// TIA Portal V20 export
FUNCTION_BLOCK "PR_UnloadingSeq_Soft2.0_workflow_f29f28"   // FB54, LAD
{ S7_Optimized_Access := 'TRUE' }
// stored: MemoryReserve 100, SetENOAutomatically false
   VAR_INPUT
      iAbort : Bool;
      iAutoRunning : Bool;
      iFaultReset : Bool;
      iGantryAtPick : Bool;
      iManualEntryConfirm : Bool;
      iPartPickOver : Bool;
      iPartPresent : Bool;
      iPickConfirmed : Bool;
      iRFIDReadError : Bool;
      iRFIDReadOver : Bool;
      iRFWriteDone : Bool;
      iRFWriteError : Bool;
      iRTR_Frm_Gantry : Bool;
      iReject : Bool;
      iReset_fault : Bool;
      iRetry : Bool;
      iRetryCount : Int;
      iSstMode : Bool;
      iSstPB : Bool;
      iStartFrmFibroSeq : Bool;
      iSystemAtHome : Bool;
      iUnloadGantryAtSafe : Bool;
   END_VAR
   VAR_OUTPUT
      qError : Array[0..2] of Bool;
      qMessage : Array[0..0] of Bool;
      qUnloadOver : Bool;
   END_VAR
   VAR
      c120_ChkPartAbsent_T1 : Bool;
      c120_ChkPartAbsent_T2 : Bool;
      c130_WtOpDecisionPick_T1 : Bool;
      c130_WtOpDecisionPick_T2 : Bool;
      c140_WtRFIDWriteOver_T1 : Bool;
      c140_WtRFIDWriteOver_T2 : Bool;
      c150_ChkRFWriteRetryCount_T1 : Bool;
      c150_ChkRFWriteRetryCount_T2 : Bool;
      c160_WtOpDecisionWrite_T1 : Bool;
      c160_WtOpDecisionWrite_T2 : Bool;
      c20_ChkRecoveryStatus_T1 : Bool;
      c20_ChkRecoveryStatus_T2 : Bool;
      c20_ChkRecoveryStatus_T3 : Bool;
      c50_WtRFIDReadOver_T1 : Bool;
      c50_WtRFIDReadOver_T2 : Bool;
      c60_ChkRetryCountOver_T1 : Bool;
      c60_ChkRetryCountOver_T2 : Bool;
      c70_WtOpDecisionRead_T1 : Bool;
      c70_WtOpDecisionRead_T2 : Bool;
      c80_ChkPartWorkable_T1 : Bool;
      c80_ChkPartWorkable_T2 : Bool;
      StateNo : Int;
      s100_WtGantryAtPick : Bool;
      s100_WtGantryAtPick_T1 : Bool;
      s10_WtStartFrmMain : Bool;
      s10_WtStartFrmMain_T1 : Bool;
      s110_WtPartPick : Bool;
      s110_WtPartPick_T1 : Bool;
      s120_ChkPartAbsent : Bool;
      s120_ChkPartAbsent_T1 : Bool;
      s120_ChkPartAbsent_T2 : Bool;
      s130_WtOpDecisionPick : Bool;
      s130_WtOpDecisionPick_T1 : Bool;
      s130_WtOpDecisionPick_T2 : Bool;
      s140_WtRFIDWriteOver : Bool;
      s140_WtRFIDWriteOver_T1 : Bool;
      s140_WtRFIDWriteOver_T2 : Bool;
      s150_ChkRFWriteRetryCount : Bool;
      s150_ChkRFWriteRetryCount_T1 : Bool;
      s150_ChkRFWriteRetryCount_T2 : Bool;
      s160_WtOpDecisionWrite : Bool;
      s160_WtOpDecisionWrite_T1 : Bool;
      s160_WtOpDecisionWrite_T2 : Bool;
      s170_ChkSystemAtHome : Bool;
      s170_ChkSystemAtHome_T1 : Bool;
      s180_WtStartLow : Bool;
      s180_WtStartLow_T1 : Bool;
      s1_WtResetReleased : Bool;
      s1_WtResetReleased_T1 : Bool;
      s20_ChkRecoveryStatus : Bool;
      s20_ChkRecoveryStatus_T1 : Bool;
      s20_ChkRecoveryStatus_T2 : Bool;
      s20_ChkRecoveryStatus_T3 : Bool;
      s30_WtOperatorAck : Bool;
      s30_WtOperatorAck_T1 : Bool;
      s40_WtAllAxesSafe : Bool;
      s40_WtAllAxesSafe_T1 : Bool;
      s50_WtRFIDReadOver : Bool;
      s50_WtRFIDReadOver_T1 : Bool;
      s50_WtRFIDReadOver_T2 : Bool;
      s60_ChkRetryCountOver : Bool;
      s60_ChkRetryCountOver_T1 : Bool;
      s60_ChkRetryCountOver_T2 : Bool;
      s70_WtOpDecisionRead : Bool;
      s70_WtOpDecisionRead_T1 : Bool;
      s70_WtOpDecisionRead_T2 : Bool;
      s80_ChkPartWorkable : Bool;
      s80_ChkPartWorkable_T1 : Bool;
      s80_ChkPartWorkable_T2 : Bool;
      s90_WtRTRFrmGantry : Bool;
      s90_WtRTRFrmGantry_T1 : Bool;
      sAbnormalStatus : Bool;
      sPartWorkable : Bool;
      sRFReadRetryCount : Int;
      sRFWriteRetryCount : Int;
      sSst : Bool;
      sSstPulse : Bool;
      sSstRise : Bool;
      sStWtResetRel : Bool;
      sStWtResetRel_T1 : Bool;
      sUnloadingActive : Bool;
   END_VAR
   VAR_TEMP
      tOne : Bool;
   END_VAR
   VAR_TEMP   // added for the SCL form of the ladder/FBD networks
      _w1 : Bool;
      _w2 : Bool;
   END_VAR
BEGIN

REGION Network 1
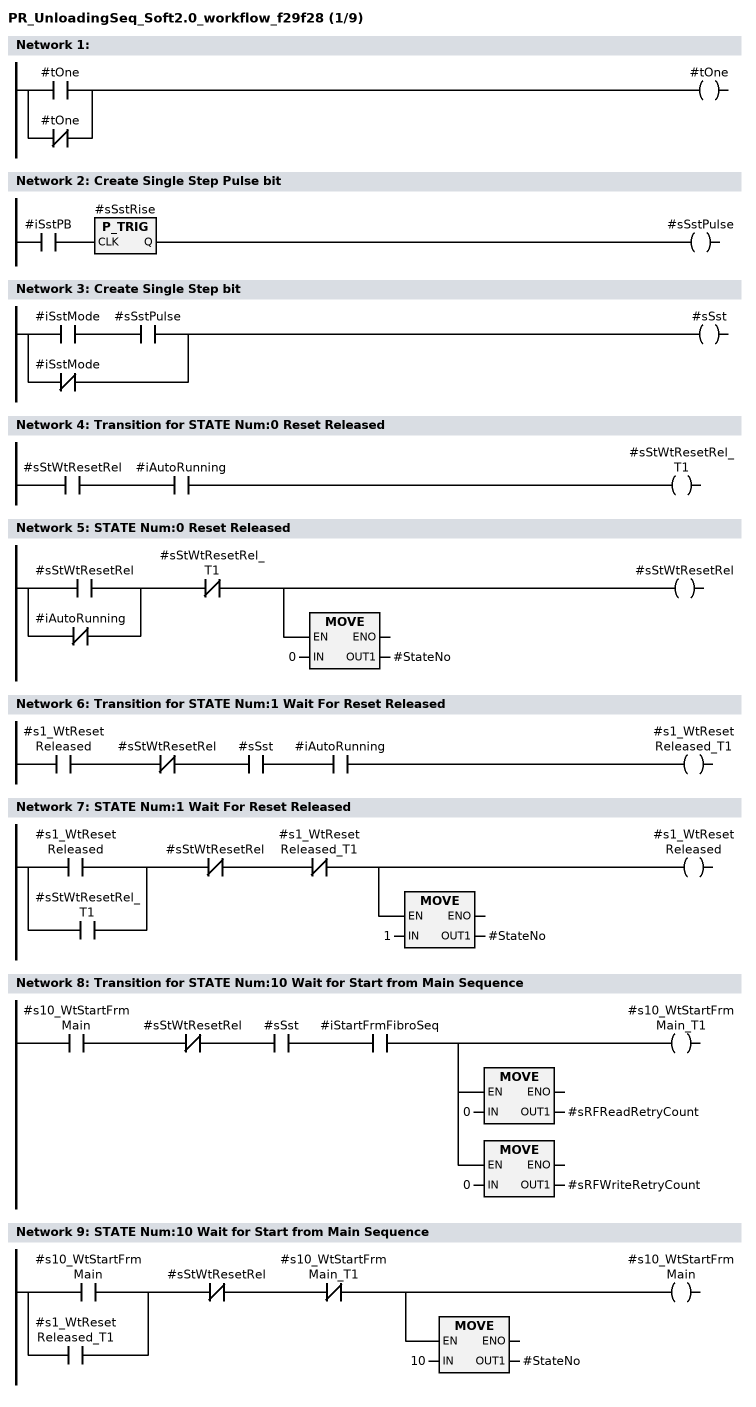
   RUNG wire#powerrail
      Contact( #tOne )
      wire#w1
      Coil( #tOne )
   END_RUNG
   RUNG wire#powerrail
      I_Contact( #tOne )
   END_RUNG wire#w1
   // the same network as SCL:
   #tOne := #tOne OR NOT #tOne;
END_REGION

REGION Network 2: Create Single Step Pulse bit
   RUNG wire#powerrail
      Contact( #iSstPB )
      P_Trig( #sSstRise )
      Coil( #sSstPulse )
   END_RUNG
   // the same network as SCL:
   #_w1 := #iSstPB AND NOT #sSstRise;   // rising edge
   #sSstRise := #iSstPB;
   #sSstPulse := #_w1;
END_REGION

REGION Network 3: Create Single Step bit
   RUNG wire#powerrail
      Contact( #iSstMode )
      Contact( #sSstPulse )
      wire#w1
      Coil( #sSst )
   END_RUNG
   RUNG wire#powerrail
      I_Contact( #iSstMode )
   END_RUNG wire#w1
   // the same network as SCL:
   #sSst := (#iSstMode AND #sSstPulse) OR NOT #iSstMode;
END_REGION

REGION Network 4: Transition for STATE Num:0 Reset Released
   RUNG wire#powerrail
      Contact( #sStWtResetRel )
      Contact( #iAutoRunning )
      Coil( #sStWtResetRel_T1 )
   END_RUNG
   // the same network as SCL:
   #sStWtResetRel_T1 := #sStWtResetRel AND #iAutoRunning;
END_REGION

REGION Network 5: STATE Num:0 Reset Released
   RUNG wire#powerrail
      Contact( #sStWtResetRel )
      wire#w1
      I_Contact( #sStWtResetRel_T1 )
      wire#w2
      Coil( #sStWtResetRel )
   END_RUNG
   RUNG wire#powerrail
      I_Contact( #iAutoRunning )
   END_RUNG wire#w1
   RUNG wire#w2
      { S7_GenerateENO := "TRUE" } Move(in := 0, out1 => #StateNo)
   END_RUNG
   // the same network as SCL:
   #sStWtResetRel := (#sStWtResetRel OR NOT #iAutoRunning) AND NOT #sStWtResetRel_T1;
   IF #sStWtResetRel THEN #StateNo := 0; END_IF;
END_REGION

REGION Network 6: Transition for STATE Num:1 Wait For Reset Released
   RUNG wire#powerrail
      Contact( #s1_WtResetReleased )
      I_Contact( #sStWtResetRel )
      Contact( #sSst )
      Contact( #iAutoRunning )
      Coil( #s1_WtResetReleased_T1 )
   END_RUNG
   // the same network as SCL:
   #s1_WtResetReleased_T1 := #s1_WtResetReleased AND NOT #sStWtResetRel AND #sSst AND #iAutoRunning;
END_REGION

REGION Network 7: STATE Num:1 Wait For Reset Released
   RUNG wire#powerrail
      Contact( #s1_WtResetReleased )
      wire#w1
      I_Contact( #sStWtResetRel )
      I_Contact( #s1_WtResetReleased_T1 )
      wire#w2
      Coil( #s1_WtResetReleased )
   END_RUNG
   RUNG wire#powerrail
      Contact( #sStWtResetRel_T1 )
   END_RUNG wire#w1
   RUNG wire#w2
      { S7_GenerateENO := "TRUE" } Move(in := 1, out1 => #StateNo)
   END_RUNG
   // the same network as SCL:
   #s1_WtResetReleased := (#s1_WtResetReleased OR #sStWtResetRel_T1) AND NOT #sStWtResetRel AND NOT #s1_WtResetReleased_T1;
   IF #s1_WtResetReleased THEN #StateNo := 1; END_IF;
END_REGION

REGION Network 8: Transition for STATE Num:10 Wait for Start from Main Sequence
   RUNG wire#powerrail
      Contact( #s10_WtStartFrmMain )
      I_Contact( #sStWtResetRel )
      Contact( #sSst )
      Contact( #iStartFrmFibroSeq )
      wire#w1
      Coil( #s10_WtStartFrmMain_T1 )
   END_RUNG
   RUNG wire#w1
      Move(in := 0, out1 => #sRFReadRetryCount)
   END_RUNG
   RUNG wire#w1
      Move(in := 0, out1 => #sRFWriteRetryCount)
   END_RUNG
   // the same network as SCL:
   #s10_WtStartFrmMain_T1 := #s10_WtStartFrmMain AND NOT #sStWtResetRel AND #sSst AND #iStartFrmFibroSeq;
   IF #s10_WtStartFrmMain_T1 THEN
       #sRFReadRetryCount := 0;
       #sRFWriteRetryCount := 0;
   END_IF;
END_REGION

REGION Network 9: STATE Num:10 Wait for Start from Main Sequence
   RUNG wire#powerrail
      Contact( #s10_WtStartFrmMain )
      wire#w1
      I_Contact( #sStWtResetRel )
      I_Contact( #s10_WtStartFrmMain_T1 )
      wire#w2
      Coil( #s10_WtStartFrmMain )
   END_RUNG
   RUNG wire#powerrail
      Contact( #s1_WtResetReleased_T1 )
   END_RUNG wire#w1
   RUNG wire#w2
      { S7_GenerateENO := "TRUE" } Move(in := 10, out1 => #StateNo)
   END_RUNG
   // the same network as SCL:
   #s10_WtStartFrmMain := (#s10_WtStartFrmMain OR #s1_WtResetReleased_T1) AND NOT #sStWtResetRel AND NOT #s10_WtStartFrmMain_T1;
   IF #s10_WtStartFrmMain THEN #StateNo := 10; END_IF;
END_REGION

REGION Network 10: Condition1 for STATE Num:20 Chek Recovery Status
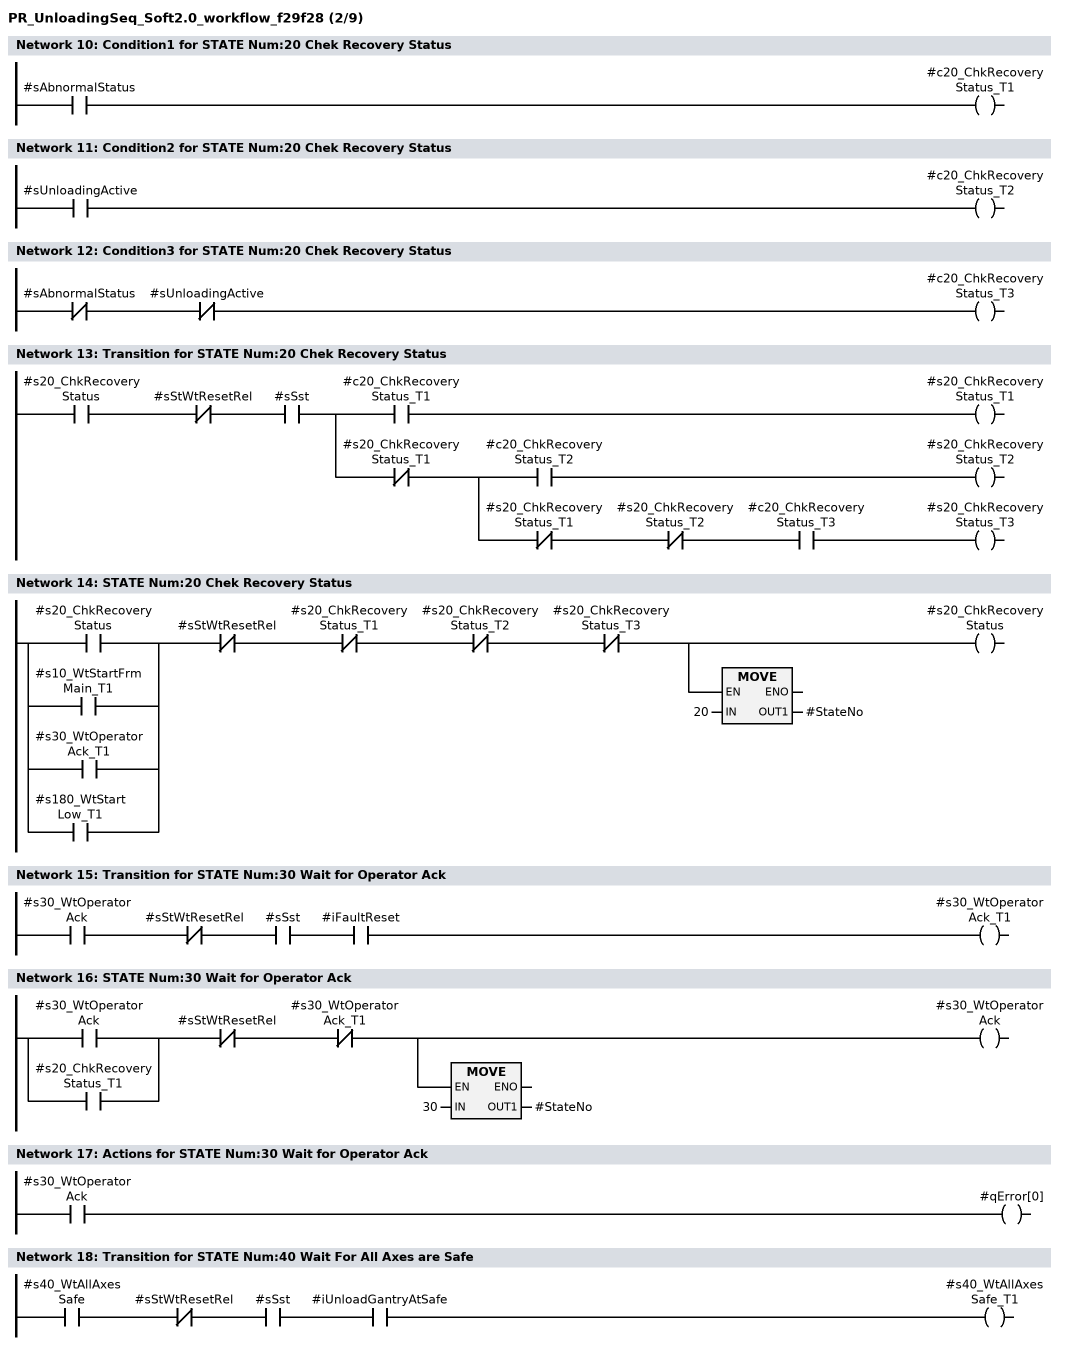
   RUNG wire#powerrail
      Contact( #sAbnormalStatus )
      Coil( #c20_ChkRecoveryStatus_T1 )
   END_RUNG
   // the same network as SCL:
   #c20_ChkRecoveryStatus_T1 := #sAbnormalStatus;
END_REGION

REGION Network 11: Condition2 for STATE Num:20 Chek Recovery Status
   RUNG wire#powerrail
      Contact( #sUnloadingActive )
      Coil( #c20_ChkRecoveryStatus_T2 )
   END_RUNG
   // the same network as SCL:
   #c20_ChkRecoveryStatus_T2 := #sUnloadingActive;
END_REGION

REGION Network 12: Condition3 for STATE Num:20 Chek Recovery Status
   RUNG wire#powerrail
      I_Contact( #sAbnormalStatus )
      I_Contact( #sUnloadingActive )
      Coil( #c20_ChkRecoveryStatus_T3 )
   END_RUNG
   // the same network as SCL:
   #c20_ChkRecoveryStatus_T3 := NOT #sAbnormalStatus AND NOT #sUnloadingActive;
END_REGION

REGION Network 13: Transition for STATE Num:20 Chek Recovery Status
   RUNG wire#powerrail
      Contact( #s20_ChkRecoveryStatus )
      I_Contact( #sStWtResetRel )
      Contact( #sSst )
      wire#w1
      Contact( #c20_ChkRecoveryStatus_T1 )
      Coil( #s20_ChkRecoveryStatus_T1 )
   END_RUNG
   RUNG wire#w1
      I_Contact( #s20_ChkRecoveryStatus_T1 )
      wire#w2
      Contact( #c20_ChkRecoveryStatus_T2 )
      Coil( #s20_ChkRecoveryStatus_T2 )
   END_RUNG
   RUNG wire#w2
      I_Contact( #s20_ChkRecoveryStatus_T1 )
      I_Contact( #s20_ChkRecoveryStatus_T2 )
      Contact( #c20_ChkRecoveryStatus_T3 )
      Coil( #s20_ChkRecoveryStatus_T3 )
   END_RUNG
   // the same network as SCL:
   #_w1 := #s20_ChkRecoveryStatus AND NOT #sStWtResetRel AND #sSst;
   #s20_ChkRecoveryStatus_T1 := #_w1 AND #c20_ChkRecoveryStatus_T1;
   #_w2 := #_w1 AND NOT #s20_ChkRecoveryStatus_T1;
   #s20_ChkRecoveryStatus_T2 := #_w2 AND #c20_ChkRecoveryStatus_T2;
   #s20_ChkRecoveryStatus_T3 := #_w2 AND NOT #s20_ChkRecoveryStatus_T1 AND NOT #s20_ChkRecoveryStatus_T2 AND #c20_ChkRecoveryStatus_T3;
END_REGION

REGION Network 14: STATE Num:20 Chek Recovery Status
   RUNG wire#powerrail
      Contact( #s20_ChkRecoveryStatus )
      wire#w1
      I_Contact( #sStWtResetRel )
      I_Contact( #s20_ChkRecoveryStatus_T1 )
      I_Contact( #s20_ChkRecoveryStatus_T2 )
      I_Contact( #s20_ChkRecoveryStatus_T3 )
      wire#w2
      Coil( #s20_ChkRecoveryStatus )
   END_RUNG
   RUNG wire#powerrail
      Contact( #s10_WtStartFrmMain_T1 )
   END_RUNG wire#w1
   RUNG wire#powerrail
      Contact( #s30_WtOperatorAck_T1 )
   END_RUNG wire#w1
   RUNG wire#powerrail
      Contact( #s180_WtStartLow_T1 )
   END_RUNG wire#w1
   RUNG wire#w2
      { S7_GenerateENO := "TRUE" } Move(in := 20, out1 => #StateNo)
   END_RUNG
   // the same network as SCL:
   #s20_ChkRecoveryStatus := (#s20_ChkRecoveryStatus OR #s10_WtStartFrmMain_T1 OR #s30_WtOperatorAck_T1 OR #s180_WtStartLow_T1) AND NOT #sStWtResetRel AND NOT #s20_ChkRecoveryStatus_T1 AND NOT #s20_ChkRecoveryStatus_T2 AND NOT #s20_ChkRecoveryStatus_T3;
   IF #s20_ChkRecoveryStatus THEN #StateNo := 20; END_IF;
END_REGION

REGION Network 15: Transition for STATE Num:30 Wait for Operator Ack
   RUNG wire#powerrail
      Contact( #s30_WtOperatorAck )
      I_Contact( #sStWtResetRel )
      Contact( #sSst )
      Contact( #iFaultReset )
      Coil( #s30_WtOperatorAck_T1 )
   END_RUNG
   // the same network as SCL:
   #s30_WtOperatorAck_T1 := #s30_WtOperatorAck AND NOT #sStWtResetRel AND #sSst AND #iFaultReset;
END_REGION

REGION Network 16: STATE Num:30 Wait for Operator Ack
   RUNG wire#powerrail
      Contact( #s30_WtOperatorAck )
      wire#w1
      I_Contact( #sStWtResetRel )
      I_Contact( #s30_WtOperatorAck_T1 )
      wire#w2
      Coil( #s30_WtOperatorAck )
   END_RUNG
   RUNG wire#powerrail
      Contact( #s20_ChkRecoveryStatus_T1 )
   END_RUNG wire#w1
   RUNG wire#w2
      { S7_GenerateENO := "TRUE" } Move(in := 30, out1 => #StateNo)
   END_RUNG
   // the same network as SCL:
   #s30_WtOperatorAck := (#s30_WtOperatorAck OR #s20_ChkRecoveryStatus_T1) AND NOT #sStWtResetRel AND NOT #s30_WtOperatorAck_T1;
   IF #s30_WtOperatorAck THEN #StateNo := 30; END_IF;
END_REGION

REGION Network 17: Actions for STATE Num:30 Wait for Operator Ack
   RUNG wire#powerrail
      Contact( #s30_WtOperatorAck )
      Coil( #qError[0] )
   END_RUNG
   // the same network as SCL:
   #qError[0] := #s30_WtOperatorAck;
END_REGION

REGION Network 18: Transition for STATE Num:40 Wait For All Axes are Safe
   RUNG wire#powerrail
      Contact( #s40_WtAllAxesSafe )
      I_Contact( #sStWtResetRel )
      Contact( #sSst )
      Contact( #iUnloadGantryAtSafe )
      Coil( #s40_WtAllAxesSafe_T1 )
   END_RUNG
   // the same network as SCL:
   #s40_WtAllAxesSafe_T1 := #s40_WtAllAxesSafe AND NOT #sStWtResetRel AND #sSst AND #iUnloadGantryAtSafe;
END_REGION

REGION Network 19: STATE Num:40 Wait For All Axes are Safe
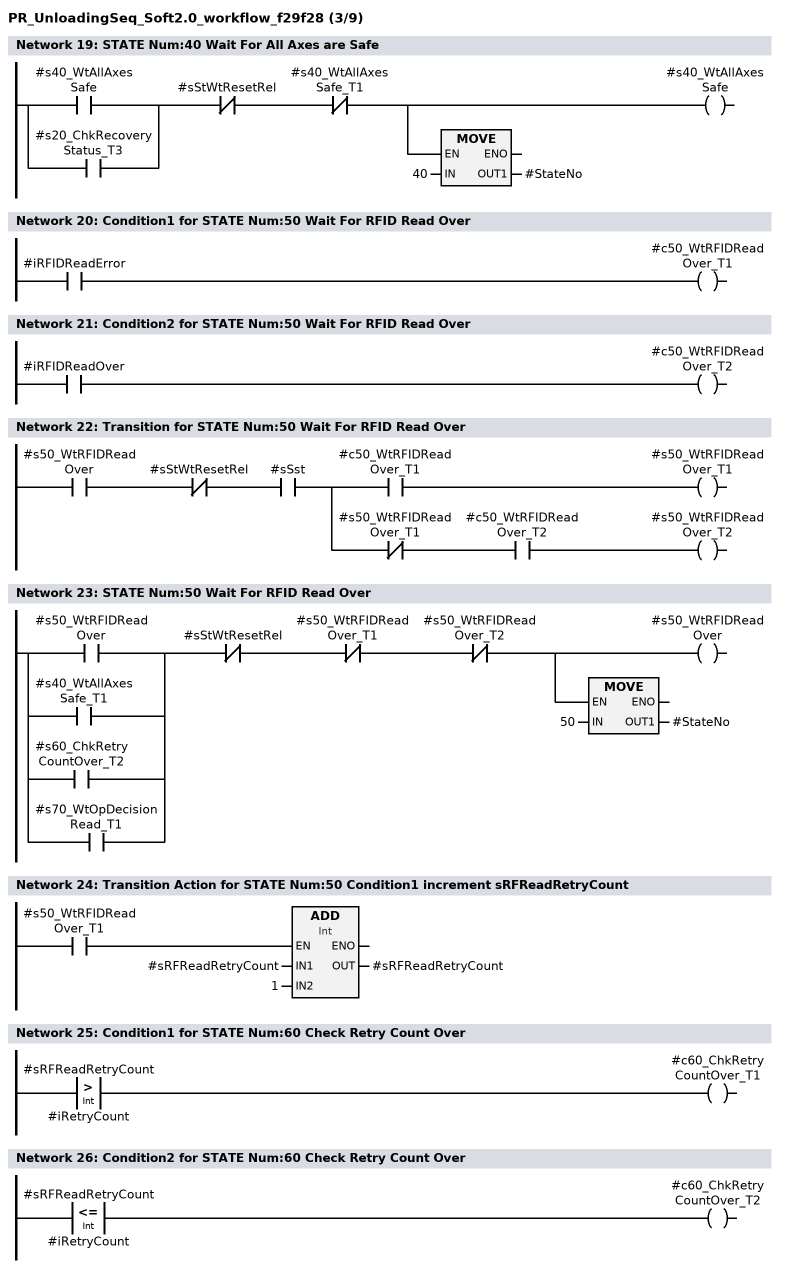
   RUNG wire#powerrail
      Contact( #s40_WtAllAxesSafe )
      wire#w1
      I_Contact( #sStWtResetRel )
      I_Contact( #s40_WtAllAxesSafe_T1 )
      wire#w2
      Coil( #s40_WtAllAxesSafe )
   END_RUNG
   RUNG wire#powerrail
      Contact( #s20_ChkRecoveryStatus_T3 )
   END_RUNG wire#w1
   RUNG wire#w2
      { S7_GenerateENO := "TRUE" } Move(in := 40, out1 => #StateNo)
   END_RUNG
   // the same network as SCL:
   #s40_WtAllAxesSafe := (#s40_WtAllAxesSafe OR #s20_ChkRecoveryStatus_T3) AND NOT #sStWtResetRel AND NOT #s40_WtAllAxesSafe_T1;
   IF #s40_WtAllAxesSafe THEN #StateNo := 40; END_IF;
END_REGION

REGION Network 20: Condition1 for STATE Num:50 Wait For RFID Read Over
   RUNG wire#powerrail
      Contact( #iRFIDReadError )
      Coil( #c50_WtRFIDReadOver_T1 )
   END_RUNG
   // the same network as SCL:
   #c50_WtRFIDReadOver_T1 := #iRFIDReadError;
END_REGION

REGION Network 21: Condition2 for STATE Num:50 Wait For RFID Read Over
   RUNG wire#powerrail
      Contact( #iRFIDReadOver )
      Coil( #c50_WtRFIDReadOver_T2 )
   END_RUNG
   // the same network as SCL:
   #c50_WtRFIDReadOver_T2 := #iRFIDReadOver;
END_REGION

REGION Network 22: Transition for STATE Num:50 Wait For RFID Read Over
   RUNG wire#powerrail
      Contact( #s50_WtRFIDReadOver )
      I_Contact( #sStWtResetRel )
      Contact( #sSst )
      wire#w1
      Contact( #c50_WtRFIDReadOver_T1 )
      Coil( #s50_WtRFIDReadOver_T1 )
   END_RUNG
   RUNG wire#w1
      I_Contact( #s50_WtRFIDReadOver_T1 )
      Contact( #c50_WtRFIDReadOver_T2 )
      Coil( #s50_WtRFIDReadOver_T2 )
   END_RUNG
   // the same network as SCL:
   #_w1 := #s50_WtRFIDReadOver AND NOT #sStWtResetRel AND #sSst;
   #s50_WtRFIDReadOver_T1 := #_w1 AND #c50_WtRFIDReadOver_T1;
   #s50_WtRFIDReadOver_T2 := #_w1 AND NOT #s50_WtRFIDReadOver_T1 AND #c50_WtRFIDReadOver_T2;
END_REGION

REGION Network 23: STATE Num:50 Wait For RFID Read Over
   RUNG wire#powerrail
      Contact( #s50_WtRFIDReadOver )
      wire#w1
      I_Contact( #sStWtResetRel )
      I_Contact( #s50_WtRFIDReadOver_T1 )
      I_Contact( #s50_WtRFIDReadOver_T2 )
      wire#w2
      Coil( #s50_WtRFIDReadOver )
   END_RUNG
   RUNG wire#powerrail
      Contact( #s40_WtAllAxesSafe_T1 )
   END_RUNG wire#w1
   RUNG wire#powerrail
      Contact( #s60_ChkRetryCountOver_T2 )
   END_RUNG wire#w1
   RUNG wire#powerrail
      Contact( #s70_WtOpDecisionRead_T1 )
   END_RUNG wire#w1
   RUNG wire#w2
      { S7_GenerateENO := "TRUE" } Move(in := 50, out1 => #StateNo)
   END_RUNG
   // the same network as SCL:
   #s50_WtRFIDReadOver := (#s50_WtRFIDReadOver OR #s40_WtAllAxesSafe_T1 OR #s60_ChkRetryCountOver_T2 OR #s70_WtOpDecisionRead_T1) AND NOT #sStWtResetRel AND NOT #s50_WtRFIDReadOver_T1 AND NOT #s50_WtRFIDReadOver_T2;
   IF #s50_WtRFIDReadOver THEN #StateNo := 50; END_IF;
END_REGION

REGION Network 24: Transition Action for STATE Num:50 Condition1 increment sRFReadRetryCount
   RUNG wire#powerrail
      Contact( #s50_WtRFIDReadOver_T1 )
      { S7_Templates := "SrcType := Int"; S7_GenerateENO := "TRUE" } Add(in1 := #sRFReadRetryCount, in2 := 1, out => #sRFReadRetryCount)
   END_RUNG
   // the same network as SCL:
   IF #s50_WtRFIDReadOver_T1 THEN #sRFReadRetryCount := #sRFReadRetryCount + 1; END_IF;
END_REGION

REGION Network 25: Condition1 for STATE Num:60 Check Retry Count Over
   RUNG wire#powerrail
      { S7_Templates := "SrcType := Int" } GT_Contact(in1 := #sRFReadRetryCount, in2 := #iRetryCount)
      Coil( #c60_ChkRetryCountOver_T1 )
   END_RUNG
   // the same network as SCL:
   #c60_ChkRetryCountOver_T1 := #sRFReadRetryCount > #iRetryCount;
END_REGION

REGION Network 26: Condition2 for STATE Num:60 Check Retry Count Over
   RUNG wire#powerrail
      { S7_Templates := "SrcType := Int" } LE_Contact(in1 := #sRFReadRetryCount, in2 := #iRetryCount)
      Coil( #c60_ChkRetryCountOver_T2 )
   END_RUNG
   // the same network as SCL:
   #c60_ChkRetryCountOver_T2 := #sRFReadRetryCount <= #iRetryCount;
END_REGION

REGION Network 27: Transition for STATE Num:60 Check Retry Count Over
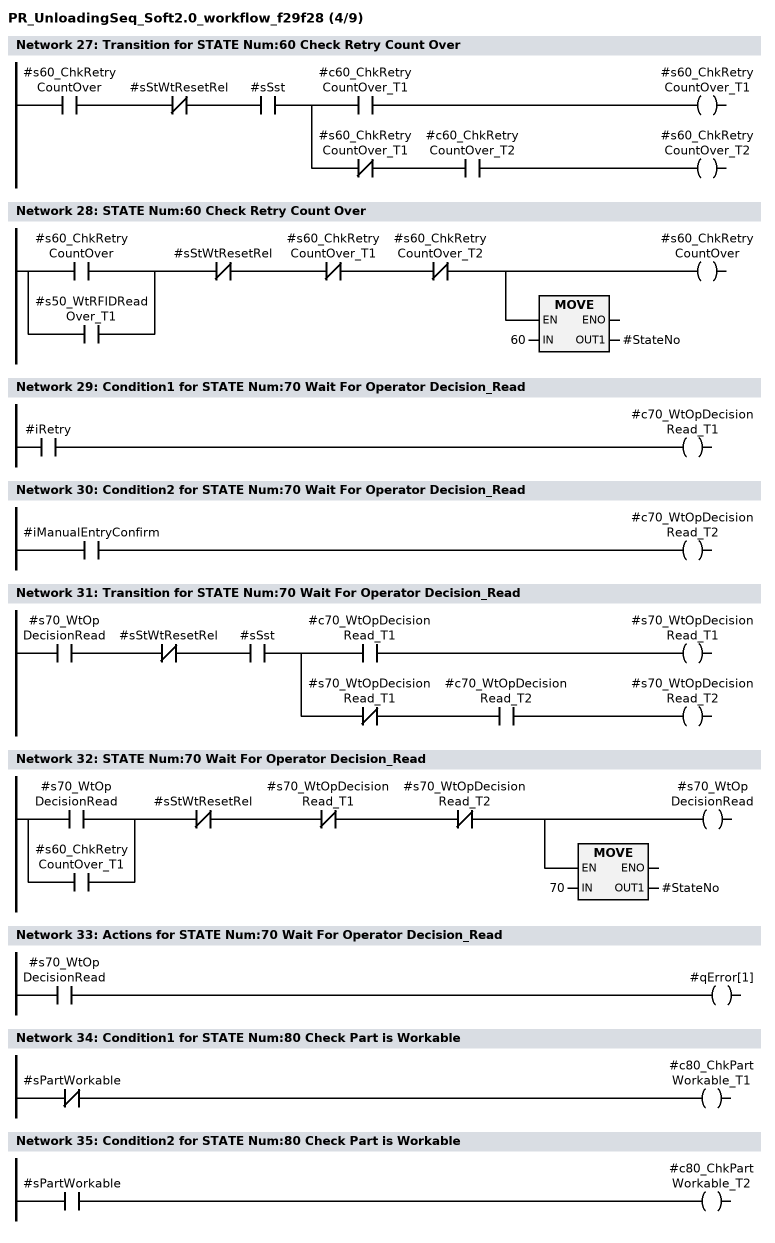
   RUNG wire#powerrail
      Contact( #s60_ChkRetryCountOver )
      I_Contact( #sStWtResetRel )
      Contact( #sSst )
      wire#w1
      Contact( #c60_ChkRetryCountOver_T1 )
      Coil( #s60_ChkRetryCountOver_T1 )
   END_RUNG
   RUNG wire#w1
      I_Contact( #s60_ChkRetryCountOver_T1 )
      Contact( #c60_ChkRetryCountOver_T2 )
      Coil( #s60_ChkRetryCountOver_T2 )
   END_RUNG
   // the same network as SCL:
   #_w1 := #s60_ChkRetryCountOver AND NOT #sStWtResetRel AND #sSst;
   #s60_ChkRetryCountOver_T1 := #_w1 AND #c60_ChkRetryCountOver_T1;
   #s60_ChkRetryCountOver_T2 := #_w1 AND NOT #s60_ChkRetryCountOver_T1 AND #c60_ChkRetryCountOver_T2;
END_REGION

REGION Network 28: STATE Num:60 Check Retry Count Over
   RUNG wire#powerrail
      Contact( #s60_ChkRetryCountOver )
      wire#w1
      I_Contact( #sStWtResetRel )
      I_Contact( #s60_ChkRetryCountOver_T1 )
      I_Contact( #s60_ChkRetryCountOver_T2 )
      wire#w2
      Coil( #s60_ChkRetryCountOver )
   END_RUNG
   RUNG wire#powerrail
      Contact( #s50_WtRFIDReadOver_T1 )
   END_RUNG wire#w1
   RUNG wire#w2
      { S7_GenerateENO := "TRUE" } Move(in := 60, out1 => #StateNo)
   END_RUNG
   // the same network as SCL:
   #s60_ChkRetryCountOver := (#s60_ChkRetryCountOver OR #s50_WtRFIDReadOver_T1) AND NOT #sStWtResetRel AND NOT #s60_ChkRetryCountOver_T1 AND NOT #s60_ChkRetryCountOver_T2;
   IF #s60_ChkRetryCountOver THEN #StateNo := 60; END_IF;
END_REGION

REGION Network 29: Condition1 for STATE Num:70 Wait For Operator Decision_Read
   RUNG wire#powerrail
      Contact( #iRetry )
      Coil( #c70_WtOpDecisionRead_T1 )
   END_RUNG
   // the same network as SCL:
   #c70_WtOpDecisionRead_T1 := #iRetry;
END_REGION

REGION Network 30: Condition2 for STATE Num:70 Wait For Operator Decision_Read
   RUNG wire#powerrail
      Contact( #iManualEntryConfirm )
      Coil( #c70_WtOpDecisionRead_T2 )
   END_RUNG
   // the same network as SCL:
   #c70_WtOpDecisionRead_T2 := #iManualEntryConfirm;
END_REGION

REGION Network 31: Transition for STATE Num:70 Wait For Operator Decision_Read
   RUNG wire#powerrail
      Contact( #s70_WtOpDecisionRead )
      I_Contact( #sStWtResetRel )
      Contact( #sSst )
      wire#w1
      Contact( #c70_WtOpDecisionRead_T1 )
      Coil( #s70_WtOpDecisionRead_T1 )
   END_RUNG
   RUNG wire#w1
      I_Contact( #s70_WtOpDecisionRead_T1 )
      Contact( #c70_WtOpDecisionRead_T2 )
      Coil( #s70_WtOpDecisionRead_T2 )
   END_RUNG
   // the same network as SCL:
   #_w1 := #s70_WtOpDecisionRead AND NOT #sStWtResetRel AND #sSst;
   #s70_WtOpDecisionRead_T1 := #_w1 AND #c70_WtOpDecisionRead_T1;
   #s70_WtOpDecisionRead_T2 := #_w1 AND NOT #s70_WtOpDecisionRead_T1 AND #c70_WtOpDecisionRead_T2;
END_REGION

REGION Network 32: STATE Num:70 Wait For Operator Decision_Read
   RUNG wire#powerrail
      Contact( #s70_WtOpDecisionRead )
      wire#w1
      I_Contact( #sStWtResetRel )
      I_Contact( #s70_WtOpDecisionRead_T1 )
      I_Contact( #s70_WtOpDecisionRead_T2 )
      wire#w2
      Coil( #s70_WtOpDecisionRead )
   END_RUNG
   RUNG wire#powerrail
      Contact( #s60_ChkRetryCountOver_T1 )
   END_RUNG wire#w1
   RUNG wire#w2
      { S7_GenerateENO := "TRUE" } Move(in := 70, out1 => #StateNo)
   END_RUNG
   // the same network as SCL:
   #s70_WtOpDecisionRead := (#s70_WtOpDecisionRead OR #s60_ChkRetryCountOver_T1) AND NOT #sStWtResetRel AND NOT #s70_WtOpDecisionRead_T1 AND NOT #s70_WtOpDecisionRead_T2;
   IF #s70_WtOpDecisionRead THEN #StateNo := 70; END_IF;
END_REGION

REGION Network 33: Actions for STATE Num:70 Wait For Operator Decision_Read
   RUNG wire#powerrail
      Contact( #s70_WtOpDecisionRead )
      Coil( #qError[1] )
   END_RUNG
   // the same network as SCL:
   #qError[1] := #s70_WtOpDecisionRead;
END_REGION

REGION Network 34: Condition1 for STATE Num:80 Check Part is Workable
   RUNG wire#powerrail
      I_Contact( #sPartWorkable )
      Coil( #c80_ChkPartWorkable_T1 )
   END_RUNG
   // the same network as SCL:
   #c80_ChkPartWorkable_T1 := NOT #sPartWorkable;
END_REGION

REGION Network 35: Condition2 for STATE Num:80 Check Part is Workable
   RUNG wire#powerrail
      Contact( #sPartWorkable )
      Coil( #c80_ChkPartWorkable_T2 )
   END_RUNG
   // the same network as SCL:
   #c80_ChkPartWorkable_T2 := #sPartWorkable;
END_REGION

REGION Network 36: Transition for STATE Num:80 Check Part is Workable
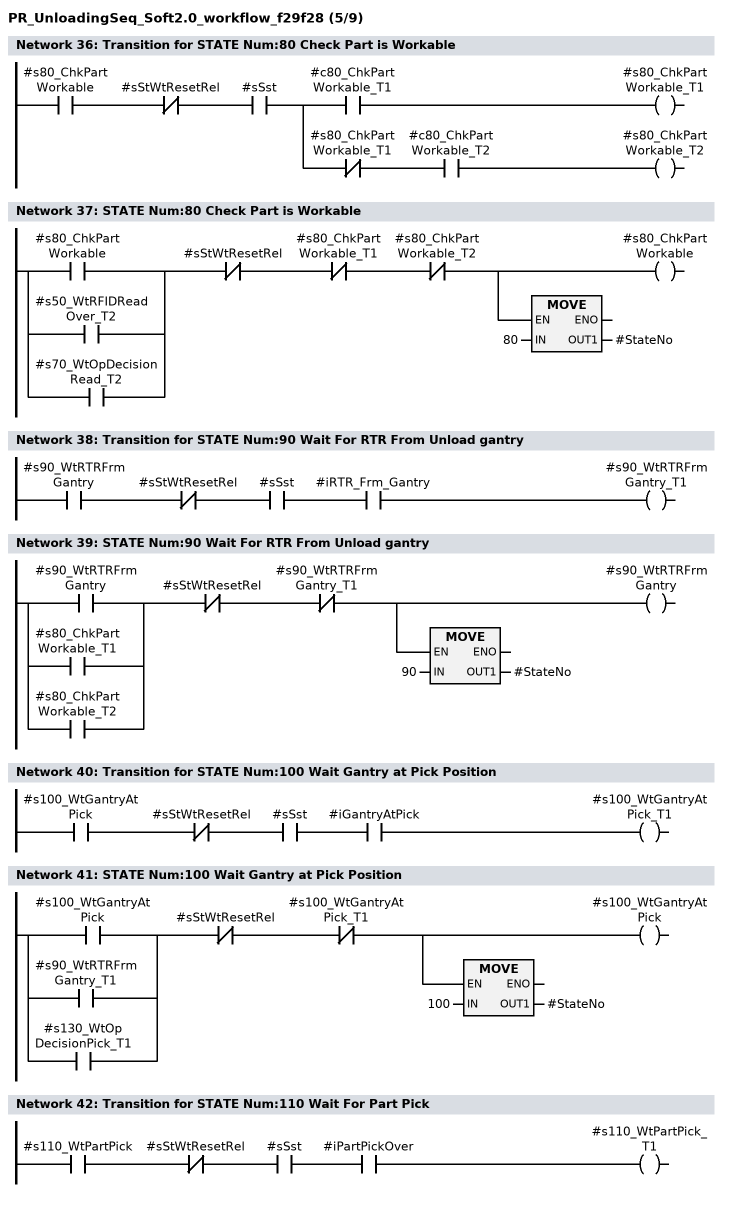
   RUNG wire#powerrail
      Contact( #s80_ChkPartWorkable )
      I_Contact( #sStWtResetRel )
      Contact( #sSst )
      wire#w1
      Contact( #c80_ChkPartWorkable_T1 )
      Coil( #s80_ChkPartWorkable_T1 )
   END_RUNG
   RUNG wire#w1
      I_Contact( #s80_ChkPartWorkable_T1 )
      Contact( #c80_ChkPartWorkable_T2 )
      Coil( #s80_ChkPartWorkable_T2 )
   END_RUNG
   // the same network as SCL:
   #_w1 := #s80_ChkPartWorkable AND NOT #sStWtResetRel AND #sSst;
   #s80_ChkPartWorkable_T1 := #_w1 AND #c80_ChkPartWorkable_T1;
   #s80_ChkPartWorkable_T2 := #_w1 AND NOT #s80_ChkPartWorkable_T1 AND #c80_ChkPartWorkable_T2;
END_REGION

REGION Network 37: STATE Num:80 Check Part is Workable
   RUNG wire#powerrail
      Contact( #s80_ChkPartWorkable )
      wire#w1
      I_Contact( #sStWtResetRel )
      I_Contact( #s80_ChkPartWorkable_T1 )
      I_Contact( #s80_ChkPartWorkable_T2 )
      wire#w2
      Coil( #s80_ChkPartWorkable )
   END_RUNG
   RUNG wire#powerrail
      Contact( #s50_WtRFIDReadOver_T2 )
   END_RUNG wire#w1
   RUNG wire#powerrail
      Contact( #s70_WtOpDecisionRead_T2 )
   END_RUNG wire#w1
   RUNG wire#w2
      { S7_GenerateENO := "TRUE" } Move(in := 80, out1 => #StateNo)
   END_RUNG
   // the same network as SCL:
   #s80_ChkPartWorkable := (#s80_ChkPartWorkable OR #s50_WtRFIDReadOver_T2 OR #s70_WtOpDecisionRead_T2) AND NOT #sStWtResetRel AND NOT #s80_ChkPartWorkable_T1 AND NOT #s80_ChkPartWorkable_T2;
   IF #s80_ChkPartWorkable THEN #StateNo := 80; END_IF;
END_REGION

REGION Network 38: Transition for STATE Num:90 Wait For RTR From Unload gantry
   RUNG wire#powerrail
      Contact( #s90_WtRTRFrmGantry )
      I_Contact( #sStWtResetRel )
      Contact( #sSst )
      Contact( #iRTR_Frm_Gantry )
      Coil( #s90_WtRTRFrmGantry_T1 )
   END_RUNG
   // the same network as SCL:
   #s90_WtRTRFrmGantry_T1 := #s90_WtRTRFrmGantry AND NOT #sStWtResetRel AND #sSst AND #iRTR_Frm_Gantry;
END_REGION

REGION Network 39: STATE Num:90 Wait For RTR From Unload gantry
   RUNG wire#powerrail
      Contact( #s90_WtRTRFrmGantry )
      wire#w1
      I_Contact( #sStWtResetRel )
      I_Contact( #s90_WtRTRFrmGantry_T1 )
      wire#w2
      Coil( #s90_WtRTRFrmGantry )
   END_RUNG
   RUNG wire#powerrail
      Contact( #s80_ChkPartWorkable_T1 )
   END_RUNG wire#w1
   RUNG wire#powerrail
      Contact( #s80_ChkPartWorkable_T2 )
   END_RUNG wire#w1
   RUNG wire#w2
      { S7_GenerateENO := "TRUE" } Move(in := 90, out1 => #StateNo)
   END_RUNG
   // the same network as SCL:
   #s90_WtRTRFrmGantry := (#s90_WtRTRFrmGantry OR #s80_ChkPartWorkable_T1 OR #s80_ChkPartWorkable_T2) AND NOT #sStWtResetRel AND NOT #s90_WtRTRFrmGantry_T1;
   IF #s90_WtRTRFrmGantry THEN #StateNo := 90; END_IF;
END_REGION

REGION Network 40: Transition for STATE Num:100 Wait Gantry at Pick Position
   RUNG wire#powerrail
      Contact( #s100_WtGantryAtPick )
      I_Contact( #sStWtResetRel )
      Contact( #sSst )
      Contact( #iGantryAtPick )
      Coil( #s100_WtGantryAtPick_T1 )
   END_RUNG
   // the same network as SCL:
   #s100_WtGantryAtPick_T1 := #s100_WtGantryAtPick AND NOT #sStWtResetRel AND #sSst AND #iGantryAtPick;
END_REGION

REGION Network 41: STATE Num:100 Wait Gantry at Pick Position
   RUNG wire#powerrail
      Contact( #s100_WtGantryAtPick )
      wire#w1
      I_Contact( #sStWtResetRel )
      I_Contact( #s100_WtGantryAtPick_T1 )
      wire#w2
      Coil( #s100_WtGantryAtPick )
   END_RUNG
   RUNG wire#powerrail
      Contact( #s90_WtRTRFrmGantry_T1 )
   END_RUNG wire#w1
   RUNG wire#powerrail
      Contact( #s130_WtOpDecisionPick_T1 )
   END_RUNG wire#w1
   RUNG wire#w2
      { S7_GenerateENO := "TRUE" } Move(in := 100, out1 => #StateNo)
   END_RUNG
   // the same network as SCL:
   #s100_WtGantryAtPick := (#s100_WtGantryAtPick OR #s90_WtRTRFrmGantry_T1 OR #s130_WtOpDecisionPick_T1) AND NOT #sStWtResetRel AND NOT #s100_WtGantryAtPick_T1;
   IF #s100_WtGantryAtPick THEN #StateNo := 100; END_IF;
END_REGION

REGION Network 42: Transition for STATE Num:110 Wait For Part Pick
   RUNG wire#powerrail
      Contact( #s110_WtPartPick )
      I_Contact( #sStWtResetRel )
      Contact( #sSst )
      Contact( #iPartPickOver )
      Coil( #s110_WtPartPick_T1 )
   END_RUNG
   // the same network as SCL:
   #s110_WtPartPick_T1 := #s110_WtPartPick AND NOT #sStWtResetRel AND #sSst AND #iPartPickOver;
END_REGION

REGION Network 43: STATE Num:110 Wait For Part Pick
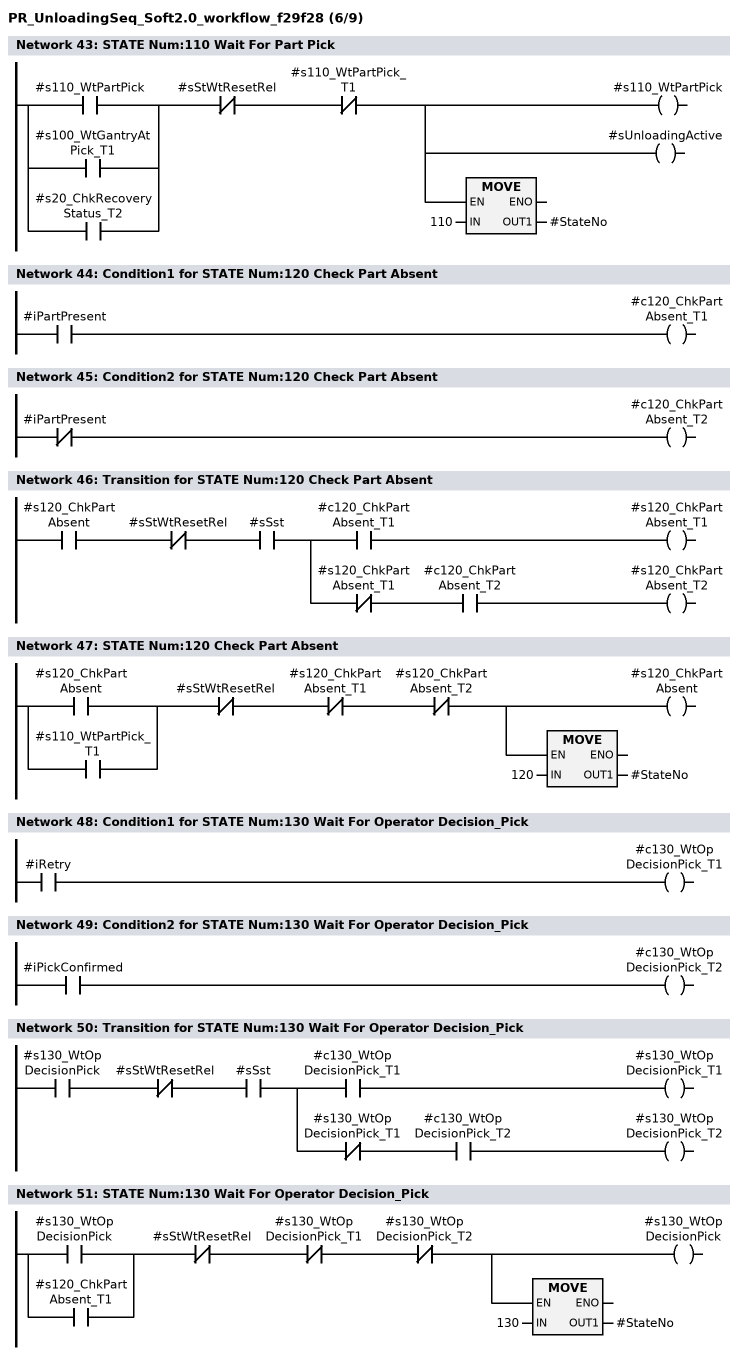
   RUNG wire#powerrail
      Contact( #s110_WtPartPick )
      wire#w1
      I_Contact( #sStWtResetRel )
      I_Contact( #s110_WtPartPick_T1 )
      wire#w2
      Coil( #s110_WtPartPick )
   END_RUNG
   RUNG wire#powerrail
      Contact( #s100_WtGantryAtPick_T1 )
   END_RUNG wire#w1
   RUNG wire#powerrail
      Contact( #s20_ChkRecoveryStatus_T2 )
   END_RUNG wire#w1
   RUNG wire#w2
      Coil( #sUnloadingActive )
   END_RUNG
   RUNG wire#w2
      { S7_GenerateENO := "TRUE" } Move(in := 110, out1 => #StateNo)
   END_RUNG
   // the same network as SCL:
   #s110_WtPartPick := (#s110_WtPartPick OR #s100_WtGantryAtPick_T1 OR #s20_ChkRecoveryStatus_T2) AND NOT #sStWtResetRel AND NOT #s110_WtPartPick_T1;
   #sUnloadingActive := #s110_WtPartPick;
   IF #s110_WtPartPick THEN #StateNo := 110; END_IF;
END_REGION

REGION Network 44: Condition1 for STATE Num:120 Check Part Absent
   RUNG wire#powerrail
      Contact( #iPartPresent )
      Coil( #c120_ChkPartAbsent_T1 )
   END_RUNG
   // the same network as SCL:
   #c120_ChkPartAbsent_T1 := #iPartPresent;
END_REGION

REGION Network 45: Condition2 for STATE Num:120 Check Part Absent
   RUNG wire#powerrail
      I_Contact( #iPartPresent )
      Coil( #c120_ChkPartAbsent_T2 )
   END_RUNG
   // the same network as SCL:
   #c120_ChkPartAbsent_T2 := NOT #iPartPresent;
END_REGION

REGION Network 46: Transition for STATE Num:120 Check Part Absent
   RUNG wire#powerrail
      Contact( #s120_ChkPartAbsent )
      I_Contact( #sStWtResetRel )
      Contact( #sSst )
      wire#w1
      Contact( #c120_ChkPartAbsent_T1 )
      Coil( #s120_ChkPartAbsent_T1 )
   END_RUNG
   RUNG wire#w1
      I_Contact( #s120_ChkPartAbsent_T1 )
      Contact( #c120_ChkPartAbsent_T2 )
      Coil( #s120_ChkPartAbsent_T2 )
   END_RUNG
   // the same network as SCL:
   #_w1 := #s120_ChkPartAbsent AND NOT #sStWtResetRel AND #sSst;
   #s120_ChkPartAbsent_T1 := #_w1 AND #c120_ChkPartAbsent_T1;
   #s120_ChkPartAbsent_T2 := #_w1 AND NOT #s120_ChkPartAbsent_T1 AND #c120_ChkPartAbsent_T2;
END_REGION

REGION Network 47: STATE Num:120 Check Part Absent
   RUNG wire#powerrail
      Contact( #s120_ChkPartAbsent )
      wire#w1
      I_Contact( #sStWtResetRel )
      I_Contact( #s120_ChkPartAbsent_T1 )
      I_Contact( #s120_ChkPartAbsent_T2 )
      wire#w2
      Coil( #s120_ChkPartAbsent )
   END_RUNG
   RUNG wire#powerrail
      Contact( #s110_WtPartPick_T1 )
   END_RUNG wire#w1
   RUNG wire#w2
      { S7_GenerateENO := "TRUE" } Move(in := 120, out1 => #StateNo)
   END_RUNG
   // the same network as SCL:
   #s120_ChkPartAbsent := (#s120_ChkPartAbsent OR #s110_WtPartPick_T1) AND NOT #sStWtResetRel AND NOT #s120_ChkPartAbsent_T1 AND NOT #s120_ChkPartAbsent_T2;
   IF #s120_ChkPartAbsent THEN #StateNo := 120; END_IF;
END_REGION

REGION Network 48: Condition1 for STATE Num:130 Wait For Operator Decision_Pick
   RUNG wire#powerrail
      Contact( #iRetry )
      Coil( #c130_WtOpDecisionPick_T1 )
   END_RUNG
   // the same network as SCL:
   #c130_WtOpDecisionPick_T1 := #iRetry;
END_REGION

REGION Network 49: Condition2 for STATE Num:130 Wait For Operator Decision_Pick
   RUNG wire#powerrail
      Contact( #iPickConfirmed )
      Coil( #c130_WtOpDecisionPick_T2 )
   END_RUNG
   // the same network as SCL:
   #c130_WtOpDecisionPick_T2 := #iPickConfirmed;
END_REGION

REGION Network 50: Transition for STATE Num:130 Wait For Operator Decision_Pick
   RUNG wire#powerrail
      Contact( #s130_WtOpDecisionPick )
      I_Contact( #sStWtResetRel )
      Contact( #sSst )
      wire#w1
      Contact( #c130_WtOpDecisionPick_T1 )
      Coil( #s130_WtOpDecisionPick_T1 )
   END_RUNG
   RUNG wire#w1
      I_Contact( #s130_WtOpDecisionPick_T1 )
      Contact( #c130_WtOpDecisionPick_T2 )
      Coil( #s130_WtOpDecisionPick_T2 )
   END_RUNG
   // the same network as SCL:
   #_w1 := #s130_WtOpDecisionPick AND NOT #sStWtResetRel AND #sSst;
   #s130_WtOpDecisionPick_T1 := #_w1 AND #c130_WtOpDecisionPick_T1;
   #s130_WtOpDecisionPick_T2 := #_w1 AND NOT #s130_WtOpDecisionPick_T1 AND #c130_WtOpDecisionPick_T2;
END_REGION

REGION Network 51: STATE Num:130 Wait For Operator Decision_Pick
   RUNG wire#powerrail
      Contact( #s130_WtOpDecisionPick )
      wire#w1
      I_Contact( #sStWtResetRel )
      I_Contact( #s130_WtOpDecisionPick_T1 )
      I_Contact( #s130_WtOpDecisionPick_T2 )
      wire#w2
      Coil( #s130_WtOpDecisionPick )
   END_RUNG
   RUNG wire#powerrail
      Contact( #s120_ChkPartAbsent_T1 )
   END_RUNG wire#w1
   RUNG wire#w2
      { S7_GenerateENO := "TRUE" } Move(in := 130, out1 => #StateNo)
   END_RUNG
   // the same network as SCL:
   #s130_WtOpDecisionPick := (#s130_WtOpDecisionPick OR #s120_ChkPartAbsent_T1) AND NOT #sStWtResetRel AND NOT #s130_WtOpDecisionPick_T1 AND NOT #s130_WtOpDecisionPick_T2;
   IF #s130_WtOpDecisionPick THEN #StateNo := 130; END_IF;
END_REGION

REGION Network 52: Condition1 for STATE Num:140 Wait for RFID Write Over
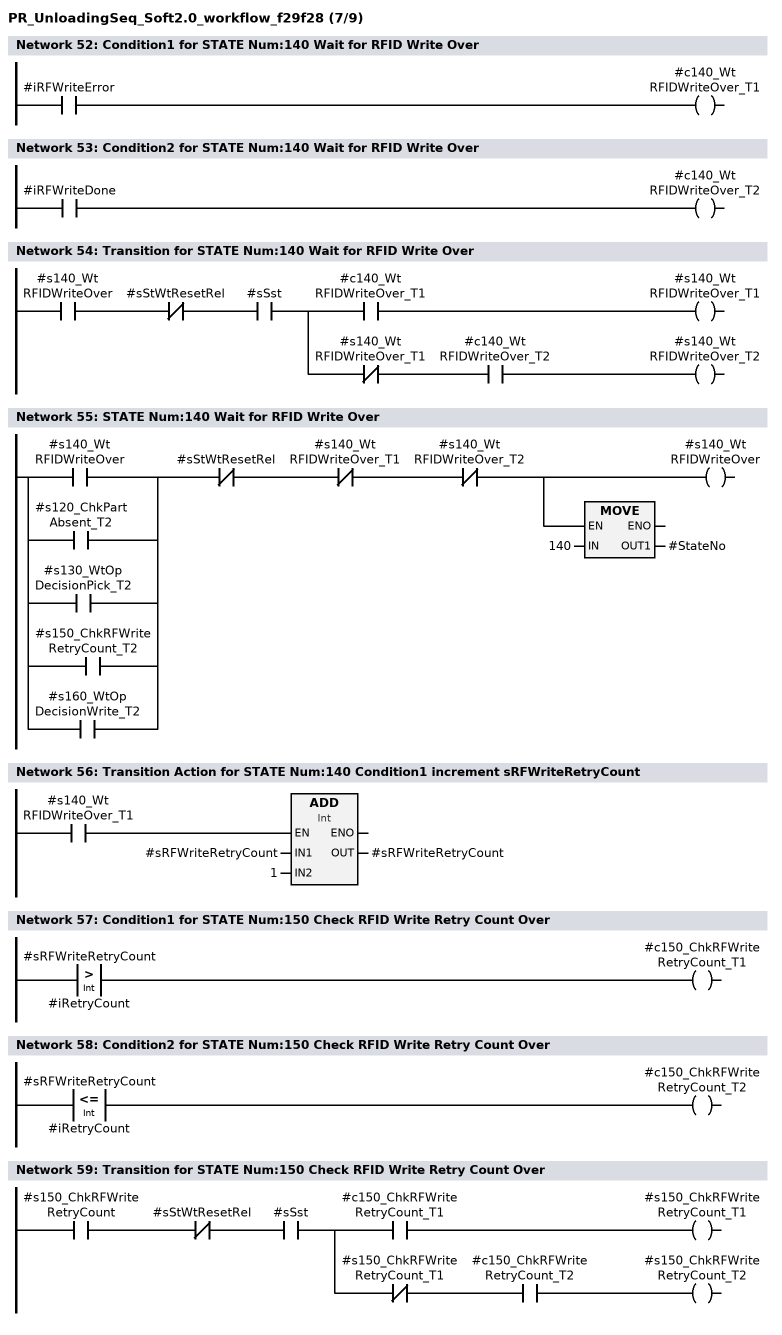
   RUNG wire#powerrail
      Contact( #iRFWriteError )
      Coil( #c140_WtRFIDWriteOver_T1 )
   END_RUNG
   // the same network as SCL:
   #c140_WtRFIDWriteOver_T1 := #iRFWriteError;
END_REGION

REGION Network 53: Condition2 for STATE Num:140 Wait for RFID Write Over
   RUNG wire#powerrail
      Contact( #iRFWriteDone )
      Coil( #c140_WtRFIDWriteOver_T2 )
   END_RUNG
   // the same network as SCL:
   #c140_WtRFIDWriteOver_T2 := #iRFWriteDone;
END_REGION

REGION Network 54: Transition for STATE Num:140 Wait for RFID Write Over
   RUNG wire#powerrail
      Contact( #s140_WtRFIDWriteOver )
      I_Contact( #sStWtResetRel )
      Contact( #sSst )
      wire#w1
      Contact( #c140_WtRFIDWriteOver_T1 )
      Coil( #s140_WtRFIDWriteOver_T1 )
   END_RUNG
   RUNG wire#w1
      I_Contact( #s140_WtRFIDWriteOver_T1 )
      Contact( #c140_WtRFIDWriteOver_T2 )
      Coil( #s140_WtRFIDWriteOver_T2 )
   END_RUNG
   // the same network as SCL:
   #_w1 := #s140_WtRFIDWriteOver AND NOT #sStWtResetRel AND #sSst;
   #s140_WtRFIDWriteOver_T1 := #_w1 AND #c140_WtRFIDWriteOver_T1;
   #s140_WtRFIDWriteOver_T2 := #_w1 AND NOT #s140_WtRFIDWriteOver_T1 AND #c140_WtRFIDWriteOver_T2;
END_REGION

REGION Network 55: STATE Num:140 Wait for RFID Write Over
   RUNG wire#powerrail
      Contact( #s140_WtRFIDWriteOver )
      wire#w1
      I_Contact( #sStWtResetRel )
      I_Contact( #s140_WtRFIDWriteOver_T1 )
      I_Contact( #s140_WtRFIDWriteOver_T2 )
      wire#w2
      Coil( #s140_WtRFIDWriteOver )
   END_RUNG
   RUNG wire#powerrail
      Contact( #s120_ChkPartAbsent_T2 )
   END_RUNG wire#w1
   RUNG wire#powerrail
      Contact( #s130_WtOpDecisionPick_T2 )
   END_RUNG wire#w1
   RUNG wire#powerrail
      Contact( #s150_ChkRFWriteRetryCount_T2 )
   END_RUNG wire#w1
   RUNG wire#powerrail
      Contact( #s160_WtOpDecisionWrite_T2 )
   END_RUNG wire#w1
   RUNG wire#w2
      { S7_GenerateENO := "TRUE" } Move(in := 140, out1 => #StateNo)
   END_RUNG
   // the same network as SCL:
   #s140_WtRFIDWriteOver := (#s140_WtRFIDWriteOver OR #s120_ChkPartAbsent_T2 OR #s130_WtOpDecisionPick_T2 OR #s150_ChkRFWriteRetryCount_T2 OR #s160_WtOpDecisionWrite_T2) AND NOT #sStWtResetRel AND NOT #s140_WtRFIDWriteOver_T1 AND NOT #s140_WtRFIDWriteOver_T2;
   IF #s140_WtRFIDWriteOver THEN #StateNo := 140; END_IF;
END_REGION

REGION Network 56: Transition Action for STATE Num:140 Condition1 increment sRFWriteRetryCount
   RUNG wire#powerrail
      Contact( #s140_WtRFIDWriteOver_T1 )
      { S7_Templates := "SrcType := Int"; S7_GenerateENO := "TRUE" } Add(in1 := #sRFWriteRetryCount, in2 := 1, out => #sRFWriteRetryCount)
   END_RUNG
   // the same network as SCL:
   IF #s140_WtRFIDWriteOver_T1 THEN #sRFWriteRetryCount := #sRFWriteRetryCount + 1; END_IF;
END_REGION

REGION Network 57: Condition1 for STATE Num:150 Check RFID Write Retry Count Over
   RUNG wire#powerrail
      { S7_Templates := "SrcType := Int" } GT_Contact(in1 := #sRFWriteRetryCount, in2 := #iRetryCount)
      Coil( #c150_ChkRFWriteRetryCount_T1 )
   END_RUNG
   // the same network as SCL:
   #c150_ChkRFWriteRetryCount_T1 := #sRFWriteRetryCount > #iRetryCount;
END_REGION

REGION Network 58: Condition2 for STATE Num:150 Check RFID Write Retry Count Over
   RUNG wire#powerrail
      { S7_Templates := "SrcType := Int" } LE_Contact(in1 := #sRFWriteRetryCount, in2 := #iRetryCount)
      Coil( #c150_ChkRFWriteRetryCount_T2 )
   END_RUNG
   // the same network as SCL:
   #c150_ChkRFWriteRetryCount_T2 := #sRFWriteRetryCount <= #iRetryCount;
END_REGION

REGION Network 59: Transition for STATE Num:150 Check RFID Write Retry Count Over
   RUNG wire#powerrail
      Contact( #s150_ChkRFWriteRetryCount )
      I_Contact( #sStWtResetRel )
      Contact( #sSst )
      wire#w1
      Contact( #c150_ChkRFWriteRetryCount_T1 )
      Coil( #s150_ChkRFWriteRetryCount_T1 )
   END_RUNG
   RUNG wire#w1
      I_Contact( #s150_ChkRFWriteRetryCount_T1 )
      Contact( #c150_ChkRFWriteRetryCount_T2 )
      Coil( #s150_ChkRFWriteRetryCount_T2 )
   END_RUNG
   // the same network as SCL:
   #_w1 := #s150_ChkRFWriteRetryCount AND NOT #sStWtResetRel AND #sSst;
   #s150_ChkRFWriteRetryCount_T1 := #_w1 AND #c150_ChkRFWriteRetryCount_T1;
   #s150_ChkRFWriteRetryCount_T2 := #_w1 AND NOT #s150_ChkRFWriteRetryCount_T1 AND #c150_ChkRFWriteRetryCount_T2;
END_REGION

REGION Network 60: STATE Num:150 Check RFID Write Retry Count Over
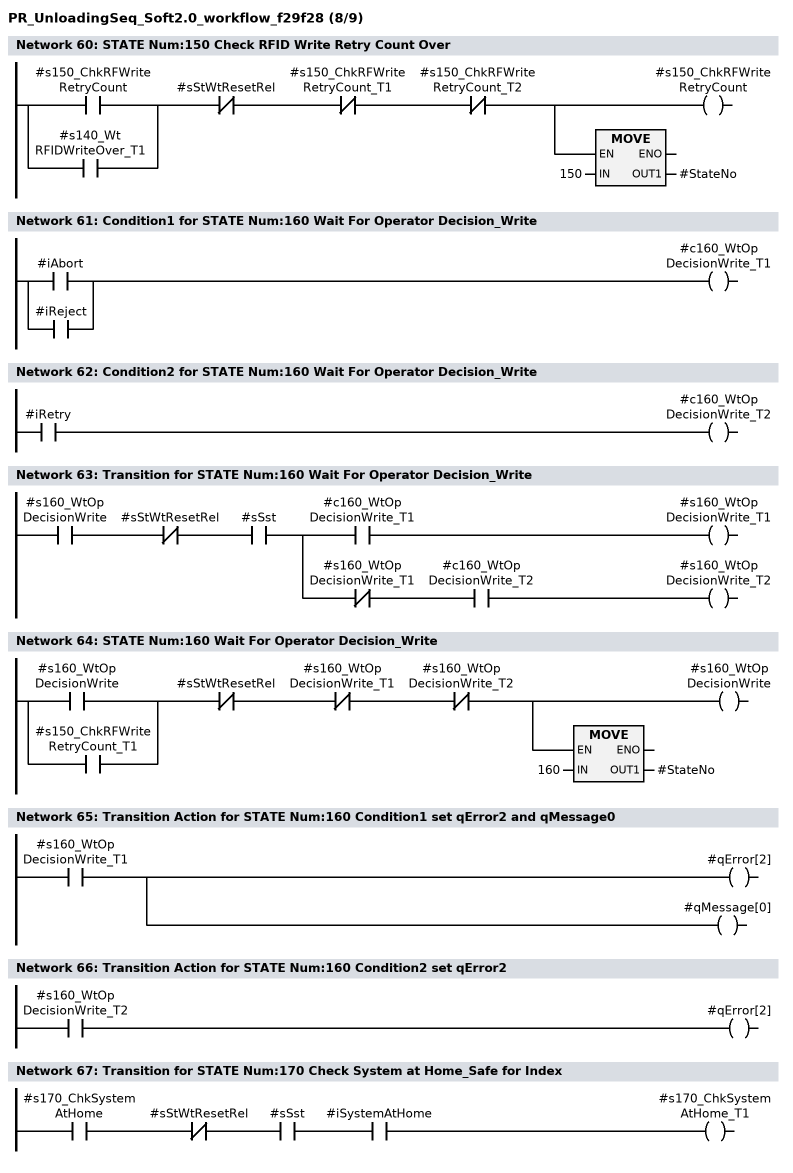
   RUNG wire#powerrail
      Contact( #s150_ChkRFWriteRetryCount )
      wire#w1
      I_Contact( #sStWtResetRel )
      I_Contact( #s150_ChkRFWriteRetryCount_T1 )
      I_Contact( #s150_ChkRFWriteRetryCount_T2 )
      wire#w2
      Coil( #s150_ChkRFWriteRetryCount )
   END_RUNG
   RUNG wire#powerrail
      Contact( #s140_WtRFIDWriteOver_T1 )
   END_RUNG wire#w1
   RUNG wire#w2
      { S7_GenerateENO := "TRUE" } Move(in := 150, out1 => #StateNo)
   END_RUNG
   // the same network as SCL:
   #s150_ChkRFWriteRetryCount := (#s150_ChkRFWriteRetryCount OR #s140_WtRFIDWriteOver_T1) AND NOT #sStWtResetRel AND NOT #s150_ChkRFWriteRetryCount_T1 AND NOT #s150_ChkRFWriteRetryCount_T2;
   IF #s150_ChkRFWriteRetryCount THEN #StateNo := 150; END_IF;
END_REGION

REGION Network 61: Condition1 for STATE Num:160 Wait For Operator Decision_Write
   RUNG wire#powerrail
      Contact( #iAbort )
      wire#w1
      Coil( #c160_WtOpDecisionWrite_T1 )
   END_RUNG
   RUNG wire#powerrail
      Contact( #iReject )
   END_RUNG wire#w1
   // the same network as SCL:
   #c160_WtOpDecisionWrite_T1 := #iAbort OR #iReject;
END_REGION

REGION Network 62: Condition2 for STATE Num:160 Wait For Operator Decision_Write
   RUNG wire#powerrail
      Contact( #iRetry )
      Coil( #c160_WtOpDecisionWrite_T2 )
   END_RUNG
   // the same network as SCL:
   #c160_WtOpDecisionWrite_T2 := #iRetry;
END_REGION

REGION Network 63: Transition for STATE Num:160 Wait For Operator Decision_Write
   RUNG wire#powerrail
      Contact( #s160_WtOpDecisionWrite )
      I_Contact( #sStWtResetRel )
      Contact( #sSst )
      wire#w1
      Contact( #c160_WtOpDecisionWrite_T1 )
      Coil( #s160_WtOpDecisionWrite_T1 )
   END_RUNG
   RUNG wire#w1
      I_Contact( #s160_WtOpDecisionWrite_T1 )
      Contact( #c160_WtOpDecisionWrite_T2 )
      Coil( #s160_WtOpDecisionWrite_T2 )
   END_RUNG
   // the same network as SCL:
   #_w1 := #s160_WtOpDecisionWrite AND NOT #sStWtResetRel AND #sSst;
   #s160_WtOpDecisionWrite_T1 := #_w1 AND #c160_WtOpDecisionWrite_T1;
   #s160_WtOpDecisionWrite_T2 := #_w1 AND NOT #s160_WtOpDecisionWrite_T1 AND #c160_WtOpDecisionWrite_T2;
END_REGION

REGION Network 64: STATE Num:160 Wait For Operator Decision_Write
   RUNG wire#powerrail
      Contact( #s160_WtOpDecisionWrite )
      wire#w1
      I_Contact( #sStWtResetRel )
      I_Contact( #s160_WtOpDecisionWrite_T1 )
      I_Contact( #s160_WtOpDecisionWrite_T2 )
      wire#w2
      Coil( #s160_WtOpDecisionWrite )
   END_RUNG
   RUNG wire#powerrail
      Contact( #s150_ChkRFWriteRetryCount_T1 )
   END_RUNG wire#w1
   RUNG wire#w2
      { S7_GenerateENO := "TRUE" } Move(in := 160, out1 => #StateNo)
   END_RUNG
   // the same network as SCL:
   #s160_WtOpDecisionWrite := (#s160_WtOpDecisionWrite OR #s150_ChkRFWriteRetryCount_T1) AND NOT #sStWtResetRel AND NOT #s160_WtOpDecisionWrite_T1 AND NOT #s160_WtOpDecisionWrite_T2;
   IF #s160_WtOpDecisionWrite THEN #StateNo := 160; END_IF;
END_REGION

REGION Network 65: Transition Action for STATE Num:160 Condition1 set qError2 and qMessage0
   RUNG wire#powerrail
      Contact( #s160_WtOpDecisionWrite_T1 )
      wire#w1
      Coil( #qError[2] )
   END_RUNG
   RUNG wire#w1
      Coil( #qMessage[0] )
   END_RUNG
   // the same network as SCL:
   #qError[2] := #s160_WtOpDecisionWrite_T1;
   #qMessage[0] := #s160_WtOpDecisionWrite_T1;
END_REGION

REGION Network 66: Transition Action for STATE Num:160 Condition2 set qError2
   RUNG wire#powerrail
      Contact( #s160_WtOpDecisionWrite_T2 )
      Coil( #qError[2] )
   END_RUNG
   // the same network as SCL:
   #qError[2] := #s160_WtOpDecisionWrite_T2;
END_REGION

REGION Network 67: Transition for STATE Num:170 Check System at Home_Safe for Index
   RUNG wire#powerrail
      Contact( #s170_ChkSystemAtHome )
      I_Contact( #sStWtResetRel )
      Contact( #sSst )
      Contact( #iSystemAtHome )
      Coil( #s170_ChkSystemAtHome_T1 )
   END_RUNG
   // the same network as SCL:
   #s170_ChkSystemAtHome_T1 := #s170_ChkSystemAtHome AND NOT #sStWtResetRel AND #sSst AND #iSystemAtHome;
END_REGION

REGION Network 68: STATE Num:170 Check System at Home_Safe for Index
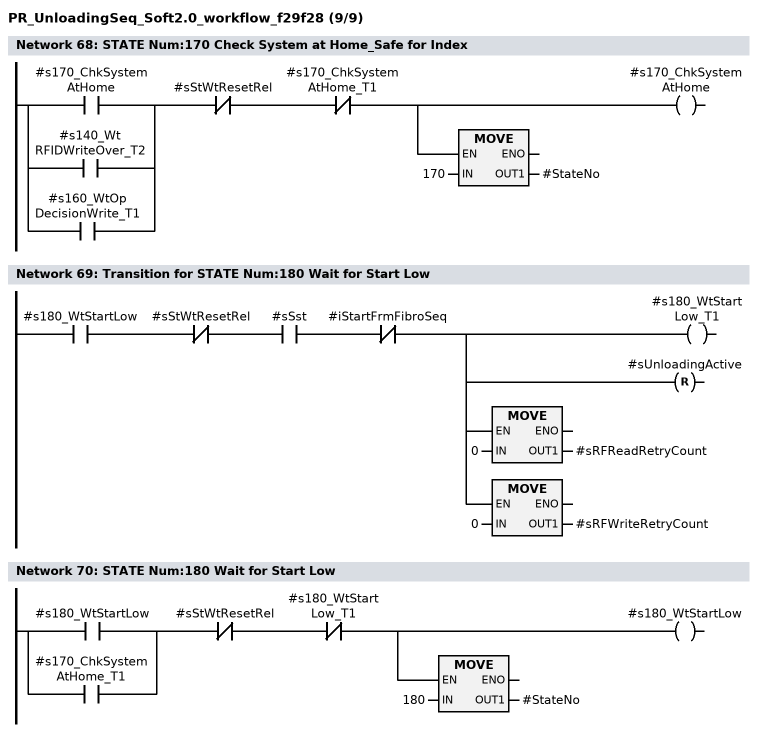
   RUNG wire#powerrail
      Contact( #s170_ChkSystemAtHome )
      wire#w1
      I_Contact( #sStWtResetRel )
      I_Contact( #s170_ChkSystemAtHome_T1 )
      wire#w2
      Coil( #s170_ChkSystemAtHome )
   END_RUNG
   RUNG wire#powerrail
      Contact( #s140_WtRFIDWriteOver_T2 )
   END_RUNG wire#w1
   RUNG wire#powerrail
      Contact( #s160_WtOpDecisionWrite_T1 )
   END_RUNG wire#w1
   RUNG wire#w2
      { S7_GenerateENO := "TRUE" } Move(in := 170, out1 => #StateNo)
   END_RUNG
   // the same network as SCL:
   #s170_ChkSystemAtHome := (#s170_ChkSystemAtHome OR #s140_WtRFIDWriteOver_T2 OR #s160_WtOpDecisionWrite_T1) AND NOT #sStWtResetRel AND NOT #s170_ChkSystemAtHome_T1;
   IF #s170_ChkSystemAtHome THEN #StateNo := 170; END_IF;
END_REGION

REGION Network 69: Transition for STATE Num:180 Wait for Start Low
   RUNG wire#powerrail
      Contact( #s180_WtStartLow )
      I_Contact( #sStWtResetRel )
      Contact( #sSst )
      I_Contact( #iStartFrmFibroSeq )
      wire#w1
      Coil( #s180_WtStartLow_T1 )
   END_RUNG
   RUNG wire#w1
      R_Coil( #sUnloadingActive )
   END_RUNG
   RUNG wire#w1
      Move(in := 0, out1 => #sRFReadRetryCount)
   END_RUNG
   RUNG wire#w1
      Move(in := 0, out1 => #sRFWriteRetryCount)
   END_RUNG
   // the same network as SCL:
   #s180_WtStartLow_T1 := #s180_WtStartLow AND NOT #sStWtResetRel AND #sSst AND NOT #iStartFrmFibroSeq;
   IF #s180_WtStartLow_T1 THEN
       #sUnloadingActive := FALSE;
       #sRFReadRetryCount := 0;
       #sRFWriteRetryCount := 0;
   END_IF;
END_REGION

REGION Network 70: STATE Num:180 Wait for Start Low
   RUNG wire#powerrail
      Contact( #s180_WtStartLow )
      wire#w1
      I_Contact( #sStWtResetRel )
      I_Contact( #s180_WtStartLow_T1 )
      wire#w2
      Coil( #s180_WtStartLow )
   END_RUNG
   RUNG wire#powerrail
      Contact( #s170_ChkSystemAtHome_T1 )
   END_RUNG wire#w1
   RUNG wire#w2
      { S7_GenerateENO := "TRUE" } Move(in := 180, out1 => #StateNo)
   END_RUNG
   // the same network as SCL:
   #s180_WtStartLow := (#s180_WtStartLow OR #s170_ChkSystemAtHome_T1) AND NOT #sStWtResetRel AND NOT #s180_WtStartLow_T1;
   IF #s180_WtStartLow THEN #StateNo := 180; END_IF;
END_REGION
END_FUNCTION_BLOCK
